// TIA Portal V21 export
// export: Created 2026-11-10T07:35:22.6089983Z, ExportSetting WithDefaults, DisplayName Totally Integrated Automation Portal, DisplayVersion V21 Update 3, DisplayName STEP 7 Professional, DisplayVersion V21 Update 3, DisplayName STEP 7 Safety, DisplayVersion V21, DisplayName Tech WebApplication, DisplayVersion V21, DisplayName WinCC Basic/Comfort/Advanced, DisplayVersion V21 Update 3, DisplayName WinCC Unified, DisplayVersion V21 Update 3
FUNCTION_BLOCK "FB_Lad_ex152"   // FB192, LAD
{ S7_Optimized_Access := 'TRUE' }
VERSION : 0.1
// stored: AutoNumber true, IsIECCheckEnabled false, IsRetainMemResEnabled false, MemoryReserve 100, SetENOAutomatically false, UDAEnableTagReadback false
   VAR_INPUT
      v_geoaddr : GEOADDR;
   END_VAR
   VAR_OUTPUT
      v_ret_val : Int;
      v_laddr : UInt;
   END_VAR
BEGIN

REGION Network 1: GEO2LOG - Determine hardware identifier from slot
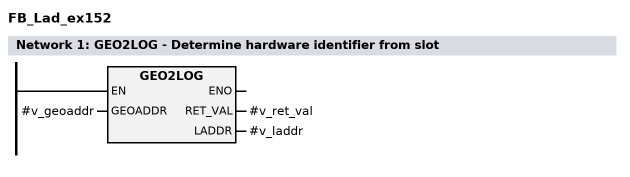
   RUNG wire#powerrail
      GEO2LOG(GEOADDR := #v_geoaddr, RET_VAL => #v_ret_val, LADDR => #v_laddr)
   END_RUNG
   // the same network as SCL:
   #v_ret_val := GEO2LOG(GEOADDR := #v_geoaddr, LADDR => #v_laddr);
END_REGION
END_FUNCTION_BLOCK
